// TIA Portal V20 export
TYPE "AZ_PrmRW_Drv2PLC"
   STRUCT
      ReadParameterID_R : Word;
      Read_WriteStatus : Struct
         "WR-END" : Bool;
         "SYS-BSY" : Bool;
         Reserved_32_bit11 : Bool;
         "WR-SET-ERR" : Bool;
         "WR-IF-ERR" : Bool;
         "WR-NV-ERR" : Bool;
         "WR-EXE-ERR" : Bool;
         "WR-ERR" : Bool;
         Reserved_33_bit0 : Bool;
         Reserved_33_bit1 : Bool;
         Reserved_33_bit2 : Bool;
         Reserved_33_bit3 : Bool;
         Reserved_33_bit4 : Bool;
         Reserved_33_bit5 : Bool;
         "RD-ERR" : Bool;
      END_STRUCT;
      WriteParameterID_R : Word;
      ReadData : DInt;
   END_STRUCT;
END_TYPE
